TYPE "ST_UnitProbeImm"
VERSION : 0.1
   STRUCT
      "Cycles" : UDInt;
      "ExitCalls" : UDInt;
      "Changes" : UDInt;
      "Resets" : UDInt;
      "AtHome" : Bool;
   END_STRUCT;
END_TYPE
